(* PLC project TBEN_L5_PLC11.project, CODESYS CODESYS V3.5 SP21 Patch 1 *)
(* stored: creationDateTime 2026-11-07T15:34:52.1459555, modificationDateTime 2026-11-07T15:09:07.4034196 *)

// Định nghĩa 1 tham số lấy từ IODD (bảng hằng trong GVL_<Model>_Def)
TYPE ST_IolParamDef :
STRUCT
    sName       : STRING(24);                  // tên theo IODD
    uiIndex     : UINT;
    usiSubindex : USINT;                       // 0 = cả index
    eType       : E_IolDataType;
    eAccess     : E_IolAccess;
    diMin       : DINT;                        // dải hợp lệ khi ghi (raw = đơn vị kỹ thuật)
    diMax       : DINT;
    diDefault   : DINT;
    sUnit       : STRING(8);
    xInReadAll  : BOOL := TRUE;                // có đọc trong ReadAll không
END_STRUCT
END_TYPE
